// TIA Portal V20 export
// export: Created 2026-10-12T05:00:29.4609343Z, ExportSetting WithDefaults, DisplayName Totally Integrated Automation Portal, DisplayVersion V20, DisplayName TIA Portal Openness, DisplayVersion V20, DisplayName TIA Portal Teamcenter Gateway, DisplayVersion V20, DisplayName TIA Portal Version Control Interface, DisplayVersion V20, DisplayName SINAMICS Startdrive Advanced, DisplayVersion V20 SP1 Update 2, DisplayName SINAMICS Startdrive G110M, G120, G120C, G120D, G120P, G115D, DisplayVersion V20 SP1 Update 2, DisplayName SINAMICS Startdrive G130, G150, S120, S150, SINAMICS MV, G220, S200, S210, DisplayVersion V20 SP1 Update 2, DisplayName STEP 7 Professional, DisplayVersion V20, DisplayName STEP 7 Safety, DisplayVersion V20, DisplayName WinCC Basic/Comfort/Advanced, DisplayVersion V20, DisplayName WinCC Professional, DisplayVersion V20, DisplayName WinCC Unified, DisplayVersion V20
FUNCTION "FRK_DecisionAudit" : Void   // FC88, SCL
{ S7_Optimized_Access := 'TRUE' }
VERSION : 0.1
// stored: AutoNumber true, IsIECCheckEnabled false, SetENOAutomatically false, UDAEnableTagReadback false
   VAR_INPUT
      Key : WString;
      SourcePath : WString;
      Option : Int;
   END_VAR
   VAR_IN_OUT
      AlarmLog : "FRK_AlarmLog";
   END_VAR
   VAR_TEMP
      Diag : "ST_Diagnostic";
      Slot : Int;
      Gone : Bool;
   END_VAR
BEGIN

   #Diag := "FRK_UnitScratch".EmptyDiagnostic;
   #Diag.Description := #Key;
   IF #Option <> 0 THEN
       #Diag.Description := CONCAT(IN1 := #Diag.Description, IN2 := WSTRING#' option=');
       #Diag.Description := CONCAT(IN1 := #Diag.Description, IN2 := STRING_TO_WSTRING(INT_TO_STRING(#Option)));
   END_IF;
   #Diag.SourcePath := #SourcePath;
   #Diag.Severity := 0;
   #Diag.Category := 0;
   #Slot := "FRK_AlarmRaise"(AlarmLog := #AlarmLog, Diag := #Diag, ResetClass := 0);
   IF #Slot > 0 THEN
       #Gone := "FRK_AlarmGone"(AlarmLog := #AlarmLog, Slot := #Slot);
   END_IF;
END_FUNCTION
